{attribute 'qualified_only'}
{attribute 'strict'}
TYPE E_BarcodeState :
(
    Idle := 0,
    Reading := 20,
    Complete := 30
);
END_TYPE

(* stored: Version 1.1.0.1
   DUT E_BarcodeState: Id {8418801c-04e1-4ce0-8b73-65aeaf094c63} *)
